(* Logix 5000 project; controller TFF vendor 1 type 14 code 107 rev 34.11; software revision 34.03; part 16 of 36 *)
(* tags used below, declared in another part *)
   Index : DINT;   // Index
   PLCDST : SINT;   // Current PLC Day Light Saving
   PLCTimeZoneString : STRING;   // Current PLC TimeZone
   TimeZoneUTC0 : STRING;   // String value for Time zone UTC 0
   Concentration : Concentration;
   ControlLoop_PCV001 : ALIAS FOR ControlLoop[3];   // PCV001 Control Loop
   ControlLoop_PCV001_5ms : ALIAS FOR ControlLoop[4];   // PCV001 Control Loop
   ControlLoop_PCV001_RAMP_OUT : REAL;   // Ramp Output
   Diafiltration : Diafiltration;
   FI101 : ALIAS FOR AnalogPoint[2];   // Filtrate Flow
   FQ_Conc : ALIAS FOR Totalizer[0];   // Concentration Totalizer
   FQ_Diaf : ALIAS FOR Totalizer[1];   // DiafiltrationTotalizer
   PCDateTime : DINT[7];   // Date/Time Array from PC
   PCV001 : ALIAS FOR AnalogPoint[3];   // Retentate Pressure Control Valve Position
   PCV001_Control : PCV_Control;   // PCV001 Control UDT
   PCV001_PID : PCV;   // PCV001 PID Management
   Phase : Phases[6];   // Phase Control Array
   PhaseTotalizer : PhaseTotalizer[18];   // Phase Totalizers Array
   Rack_Murr_Node1_TF2S : IO_Station;   // Status of Node 1 TF2S
   Rack_Murr_Node1_TF3S : IO_Station;   // Status of Node 1 TF3S
   RawAnalogInputArray : INT[50];   // Array of analog input raw
   SysControl : SysControl;   // General system status and command
   ThisSystem : SystemType;
   TimerControl : TimerControl;   // Timer Control
   Timers : Timers[22];   // Timer Array
   Totalizer : Totalizers[20];   // Totalizers Array
   Valve : Valve[100];   // Valve Array
(* MainProgram, continued *)

ROUTINE modTotal   (* ladder *)
// Totalizer Module
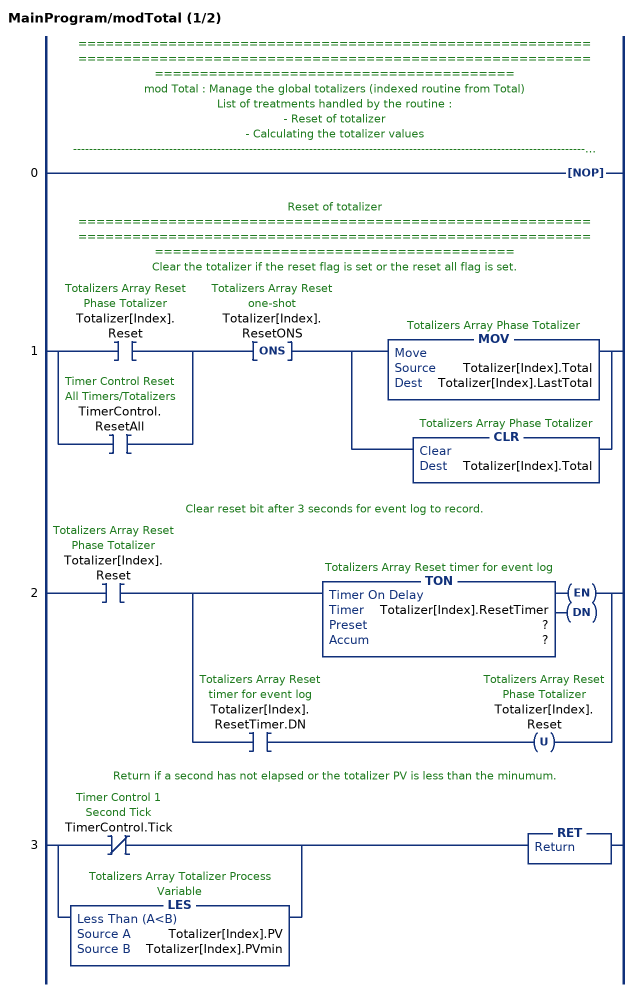
   // ==========================================================================================================================================================
   //                                                                                                   mod Total : Manage the global totalizers (indexed routine from Total)
   //                                                     List of treatments handled by the routine :
   //                                                          - Reset of totalizer
   //                                                          - Calculating the totalizer values
   //                                                     -----------------------------------------------------------------------------------------------------------------------------------------------------
   //                                                     History
   //                                                         2019-AUG-13 - Actemium - B. Roch - Initial version for Candidate Release 3.00.00.00.a
   // ==========================================================================================================================================================
   0: NOP();
   // Reset of totalizer
   // ==========================================================================================================================================================
   // Clear the totalizer if the reset flag is set or the reset all flag is set.
   1: [XIC(Totalizer[Index].Reset) ,XIC(TimerControl.ResetAll) ]ONS(Totalizer[Index].ResetONS)[MOV(Totalizer[Index].Total,Totalizer[Index].LastTotal) ,CLR(Totalizer[Index].Total) ];
   // Clear reset bit after 3 seconds for event log to record.
   2: XIC(Totalizer[Index].Reset)[TON(Totalizer[Index].ResetTimer,?,?) ,XIC(Totalizer[Index].ResetTimer.DN) OTU(Totalizer[Index].Reset) ];
   // Return if a second has not elapsed or the totalizer PV is less than the minumum.
   3: [XIO(TimerControl.Tick) ,LES(Totalizer[Index].PV,Totalizer[Index].PVmin) ]RET();
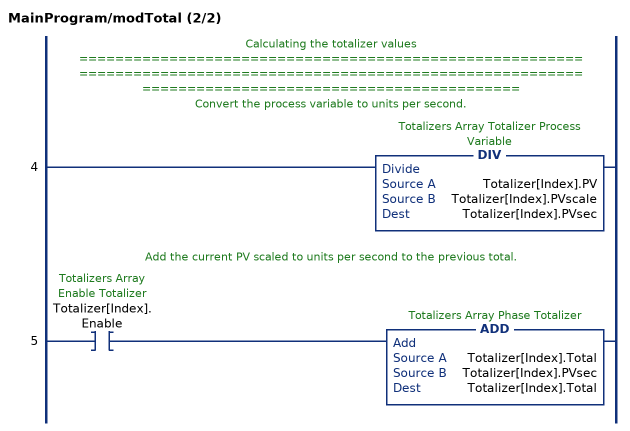
   // Calculating the totalizer values
   // ==========================================================================================================================================================
   // Convert the process variable to units per second.
   4: DIV(Totalizer[Index].PV,Totalizer[Index].PVscale,Totalizer[Index].PVsec);
   // Add the current PV scaled to units per second to the previous total.
   5: XIC(Totalizer[Index].Enable)ADD(Totalizer[Index].Total,Totalizer[Index].PVsec,Totalizer[Index].Total);
END_ROUTINE

ROUTINE PCDateTime   (* structured text *)
   (* =======================================================================
   	PCDateTime : Synchronize the PLC with PC clock
   
   	List of treatments
   		- Synchronization
   
   -----------------------------------------------------------------------------------------------------------------------------------------------------
   	History
   		2019-AUG-13 - ACTEMIUM - B. Roch - Initial version for Candidate Release 3.00.00.00.a
   		2020-SEP-14 - MERCK - Q. Spindler - Modifications for Candidate Release 3.00.00.01.a
   					- Add PLC TimeZone and DST forced settings
   =========================================================================*)
   
   
   (* Synchronization
   =========================================================================*)
   (*Update the internal PLC clock with the PC clock when the microseconds value is not -1*)
   IF PCDateTime[6] <> -1 THEN;
   	SSV (WALLCLOCKTIME, , DateTime, PCDateTime[0]);
   	PCDateTime[6] := -1;
   END_IF;
   
   (*Get PLC DST settings and set it to 0 of not already*)
   GSV (WALLCLOCKTIME, ,ApplyDST , PLCDST);
   IF PLCDST <> 0 THEN;
   	PLCDST := 0;
   	SSV (WALLCLOCKTIME, ,ApplyDST , PLCDST);
   END_IF;
   
   (*Get PLC TimeZone and set it to UTC0 of not already*)
   GSV (WALLCLOCKTIME, ,TimeZoneString, PLCTimeZoneString);
   IF PLCTimeZoneString <> TimeZoneUTC0 THEN;
   	SSV (WALLCLOCKTIME, ,TimeZoneString , TimeZoneUTC0);
   END_IF;
   
END_ROUTINE

ROUTINE Time   (* ladder *)
// Timekeeping Routine
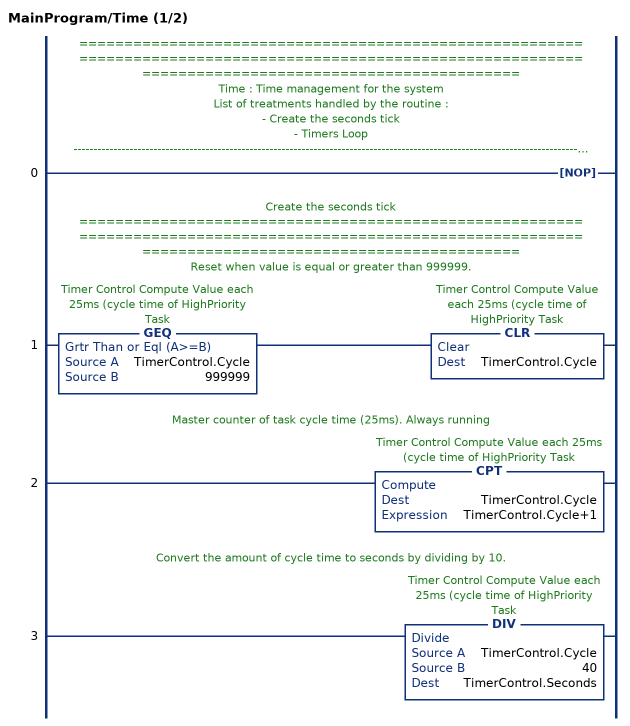
   // ==========================================================================================================================================================
   //                                                                                                                       Time : Time management for the system
   //                                                     List of treatments handled by the routine :
   //                                                          - Create the seconds tick
   //                                                          - Timers Loop
   //                                                     -----------------------------------------------------------------------------------------------------------------------------------------------------
   //                                                     History
   //                                                          2019-AUG-13 - Actemium - B. Roch - Initial version for Candidate Release 3.00.00.00.a
   //                                                          2020-SEP-14 - Merck - Q. Spindler - Modifications for Candidate Release 3.00.00.01.a
   //                                                                  - Add TimerControl.NewTickMainTask for 1 sec tick in Main task
   // ==========================================================================================================================================================
   0: NOP();
   // Create the seconds tick
   // ==========================================================================================================================================================
   // Reset when value is equal or greater than 999999.
   1: GEQ(TimerControl.Cycle,999999)CLR(TimerControl.Cycle);
   // Master counter of task cycle time (25ms). Always running
   2: CPT(TimerControl.Cycle,TimerControl.Cycle+1);
   // Convert the amount of cycle time to seconds by dividing by 10.
   3: DIV(TimerControl.Cycle,40,TimerControl.Seconds);
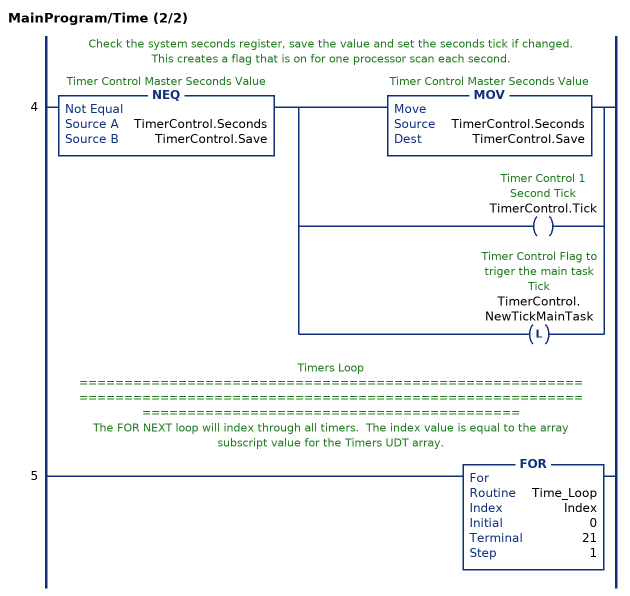
   // Check the system seconds register, save the value and set the seconds tick if changed.  This creates a flag that is on for one processor scan each second.
   4: NEQ(TimerControl.Seconds,TimerControl.Save)[MOV(TimerControl.Seconds,TimerControl.Save) ,OTE(TimerControl.Tick) ,OTL(TimerControl.NewTickMainTask) ];
   // Timers Loop
   // ==========================================================================================================================================================
   // The FOR NEXT loop will index through all timers.  The index value is equal to the array subscript value for the Timers UDT array.
   5: FOR(Time_Loop,Index,0,21,1);
END_ROUTINE

ROUTINE Time_Loop   (* ladder *)
// Timer Routine
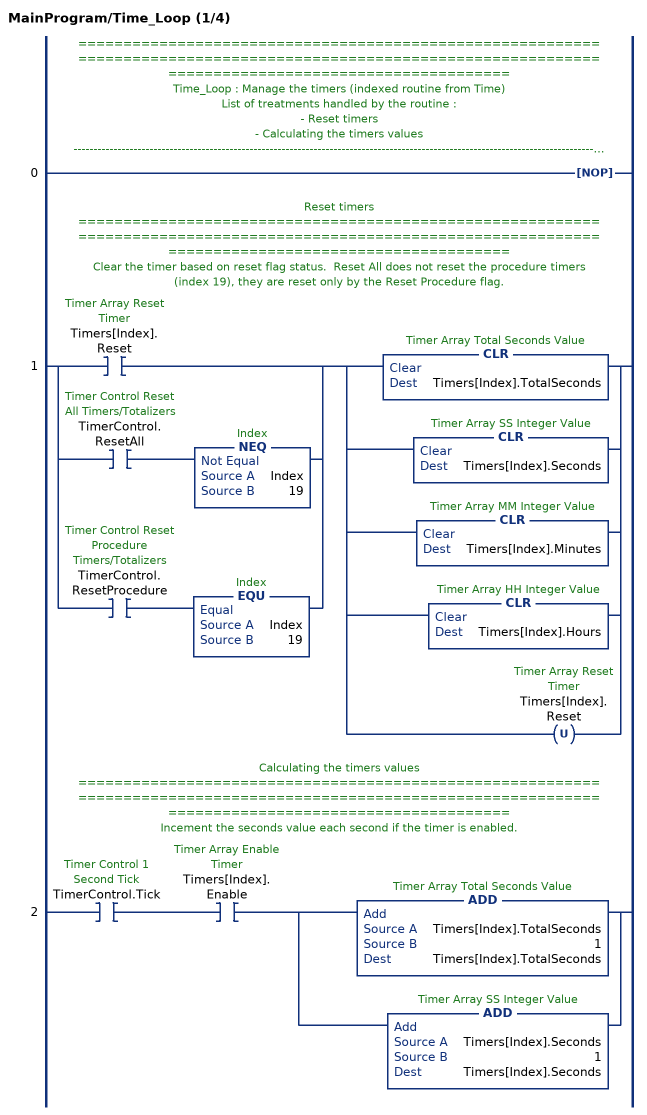
   // ==========================================================================================================================================================
   //                                                                                                              Time_Loop : Manage the timers (indexed routine from Time)
   //                                                     List of treatments handled by the routine :
   //                                                          - Reset timers
   //                                                          - Calculating the timers values
   //                                                     -----------------------------------------------------------------------------------------------------------------------------------------------------
   //                                                     History
   //                                                         2019-AUG-13 - Actemium - B. Roch - Initial version for Candidate Release 3.00.00.00.a
   // ==========================================================================================================================================================
   0: NOP();
   // Reset timers
   // ==========================================================================================================================================================
   // Clear the timer based on reset flag status.  Reset All does not reset the procedure timers (index 19), they are reset only by the Reset Procedure flag.
   1: [XIC(Timers[Index].Reset) ,XIC(TimerControl.ResetAll) NEQ(Index,19) ,XIC(TimerControl.ResetProcedure) EQU(Index,19) ][CLR(Timers[Index].TotalSeconds) ,CLR(Timers[Index].Seconds) ,CLR(Timers[Index].Minutes) ,CLR(Timers[Index].Hours) ,OTU(Timers[Index].Reset) ];
   // Calculating the timers values
   // ==========================================================================================================================================================
   // Incement the seconds value each second if the timer is enabled.
   2: XIC(TimerControl.Tick)XIC(Timers[Index].Enable)[ADD(Timers[Index].TotalSeconds,1,Timers[Index].TotalSeconds) ,ADD(Timers[Index].Seconds,1,Timers[Index].Seconds) ];
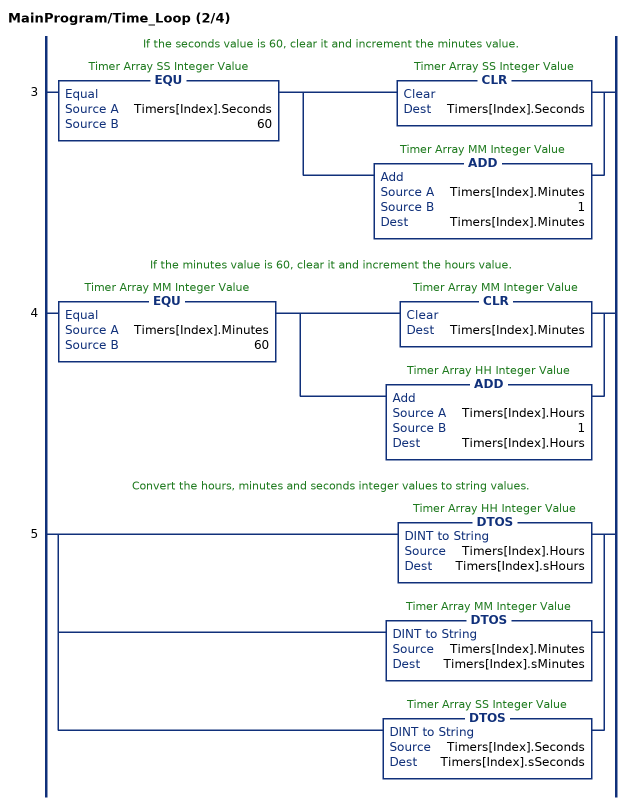
   // If the seconds value is 60, clear it and increment the minutes value.
   3: EQU(Timers[Index].Seconds,60)[CLR(Timers[Index].Seconds) ,ADD(Timers[Index].Minutes,1,Timers[Index].Minutes) ];
   // If the minutes value is 60, clear it and increment the hours value.
   4: EQU(Timers[Index].Minutes,60)[CLR(Timers[Index].Minutes) ,ADD(Timers[Index].Hours,1,Timers[Index].Hours) ];
   // Convert the hours, minutes and seconds integer values to string values.
   5: [DTOS(Timers[Index].Hours,Timers[Index].sHours) ,DTOS(Timers[Index].Minutes,Timers[Index].sMinutes) ,DTOS(Timers[Index].Seconds,Timers[Index].sSeconds) ];
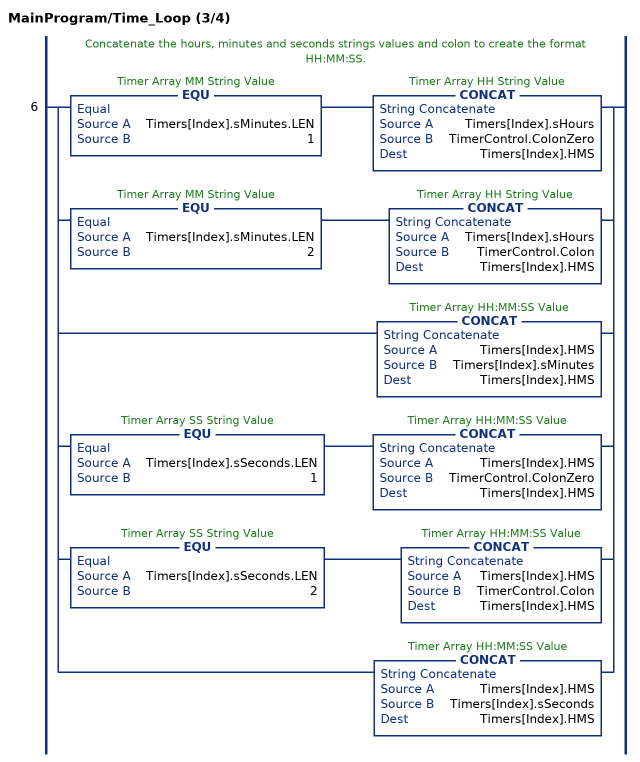
   // Concatenate the hours, minutes and seconds strings values and colon to create the format HH:MM:SS.
   6: [EQU(Timers[Index].sMinutes.LEN,1) CONCAT(Timers[Index].sHours,TimerControl.ColonZero,Timers[Index].HMS) ,EQU(Timers[Index].sMinutes.LEN,2) CONCAT(Timers[Index].sHours,TimerControl.Colon,Timers[Index].HMS) ,CONCAT(Timers[Index].HMS,Timers[Index].sMinutes,Timers[Index].HMS) ,EQU(Timers[Index].sSeconds.LEN,1) CONCAT(Timers[Index].HMS,TimerControl.ColonZero,Timers[Index].HMS) ,EQU(Timers[Index].sSeconds.LEN,2) CONCAT(Timers[Index].HMS,TimerControl.Colon,Timers[Index].HMS) ,CONCAT(Timers[Index].HMS,Timers[Index].sSeconds,Timers[Index].HMS) ];
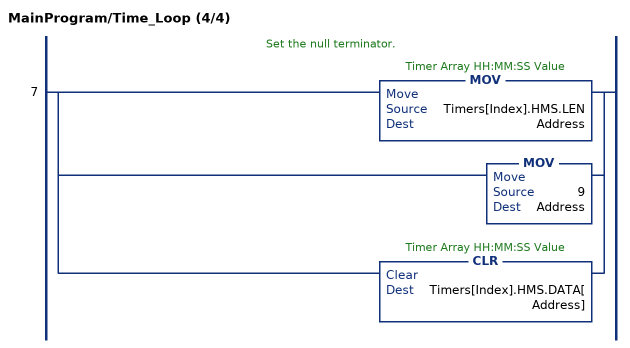
   // Set the null terminator.
   7: [[MOV(Timers[Index].HMS.LEN,Address) ,MOV(9,Address) ] ,CLR(Timers[Index].HMS.DATA[Address]) ];
END_ROUTINE

ROUTINE Total   (* ladder *)
// Totalizer Routine
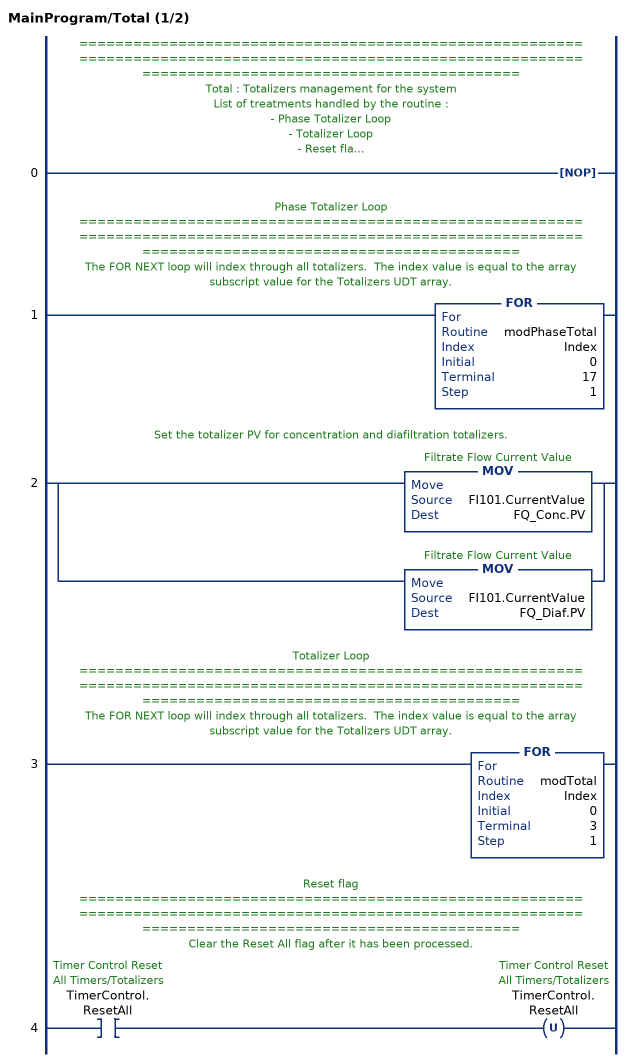
   // ==========================================================================================================================================================
   //                                                                                                              Total : Totalizers management for the system
   //                                                     List of treatments handled by the routine :
   //                                                          - Phase Totalizer Loop
   //                                                          - Totalizer Loop
   //                                                          - Reset flag
   //                                                     -----------------------------------------------------------------------------------------------------------------------------------------------------
   //                                                     History
   //                                                          2019-AUG-13 - Actemium - B. Roch - Initial version for Candidate Release 3.00.00.00.a
   // 		2020-SEP-29 - Merck - Q. Spindler - Modifications for Candidate Release 3.00.00.01.a
   // 							- Change array size of PhaseTotalizer
   // ==========================================================================================================================================================
   0: NOP();
   // Phase Totalizer Loop
   // ==========================================================================================================================================================
   // The FOR NEXT loop will index through all totalizers.  The index value is equal to the array subscript value for the Totalizers UDT array.
   1: FOR(modPhaseTotal,Index,0,17,1);
   // Set the totalizer PV for concentration and diafiltration totalizers.
   2: [MOV(FI101.CurrentValue,FQ_Conc.PV) ,MOV(FI101.CurrentValue,FQ_Diaf.PV) ];
   // Totalizer Loop
   // ==========================================================================================================================================================
   // The FOR NEXT loop will index through all totalizers.  The index value is equal to the array subscript value for the Totalizers UDT array.
   3: FOR(modTotal,Index,0,3,1);
   // Reset flag
   // ==========================================================================================================================================================
   // Clear the Reset All flag after it has been processed.
   4: XIC(TimerControl.ResetAll)OTU(TimerControl.ResetAll);
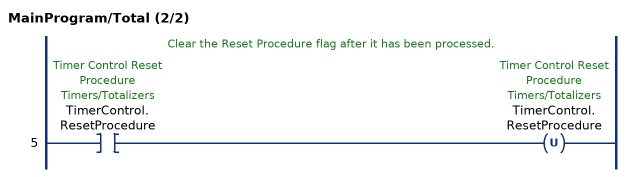
   // Clear the Reset Procedure flag after it has been processed.
   5: XIC(TimerControl.ResetProcedure)OTU(TimerControl.ResetProcedure);
END_ROUTINE
END_PROGRAM

PROGRAM MainProgram5ms   (* main routine MainRoutine, fault routine FaultRoutine *)
VAR
   Address : DINT := 1;   // Index
   Address2 : DINT := 41;
   ONS_PID02 : BOOL;
   PCV001_PID_Settings : INT;
   PCV101_PID_Settings : INT;
   SCL : SCALE := (InRawMax := 99999.0, InEUMax := 999.99);   // Scale Function
END_VAR

ROUTINE Control_Loop_PCV001_5ms   (* ladder *)
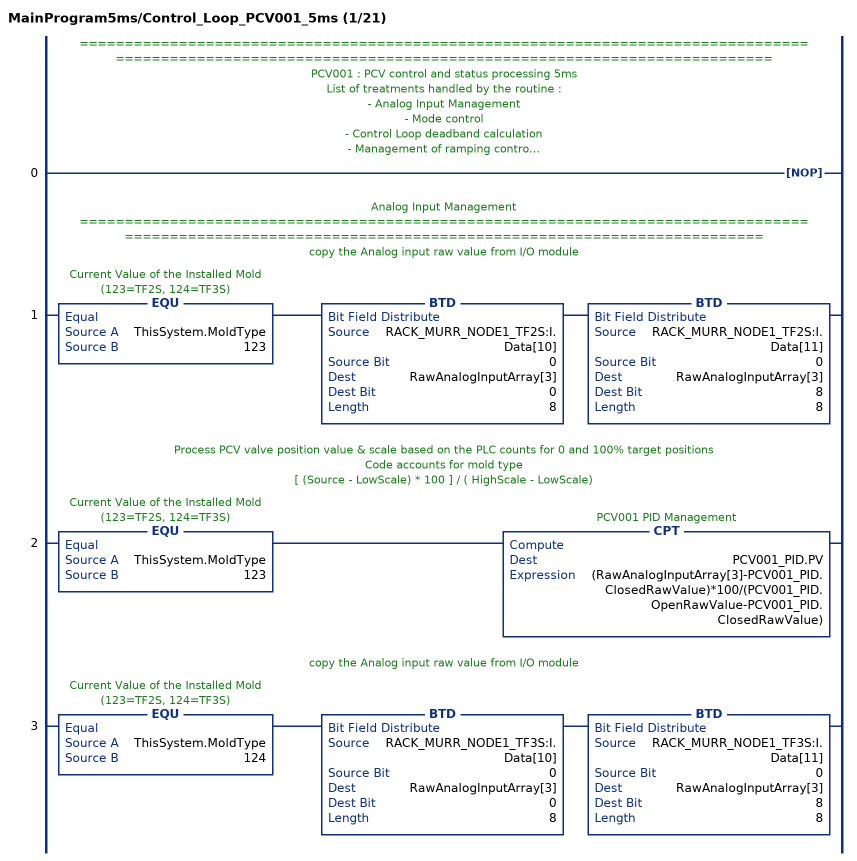
   // ==========================================================================================================================================================
   //                                                  PCV001 : PCV control and status processing 5ms
   //                                                     List of treatments handled by the routine :
   //                                                          - Analog Input Management
   //                                                          - Mode control
   //                                                          - Control Loop deadband calculation
   //                                                          - Management of ramping control
   //                                                          - Management of PID instruction
   //                                                          - PCV001 Control Valve Calibration
   //                                                          - Control of the analog output
   //                                                          - Loop status for HMI
   //                                                     -----------------------------------------------------------------------------------------------------------------------------------------------------
   //                                                     History
   //                                                          2019-AUG-13 - Actemium - B. Roch - Initial version for Candidate Release 3.00.00.00.a
   // 		                                2019-SEP-26 - ACTEMIUM - B. Roch - Modifications for Candidate Release 3.00.00.00.c
   // 					- Change compute for Analog Input Managment
   //                                                                                - Update Ramping up and down conditions
   // ==========================================================================================================================================================
   0: NOP();
   // Analog Input Management
   // ========================================================================================================================================================
   // copy the Analog input raw value from I/O module
   1: EQU(ThisSystem.MoldType,123)BTD(RACK_MURR_NODE1_TF2S:I.Data[10],0,RawAnalogInputArray[3],0,8)BTD(RACK_MURR_NODE1_TF2S:I.Data[11],0,RawAnalogInputArray[3],8,8);
   // Process PCV valve position value & scale based on the PLC counts for 0 and 100% target positions
   // Code accounts for mold type
   // [ (Source - LowScale) * 100 ] / ( HighScale - LowScale)
   2: EQU(ThisSystem.MoldType,123)CPT(PCV001_PID.PV,(RawAnalogInputArray[3]-PCV001_PID.ClosedRawValue)*100/(PCV001_PID.OpenRawValue-PCV001_PID.ClosedRawValue));
   // copy the Analog input raw value from I/O module
   3: EQU(ThisSystem.MoldType,124)BTD(RACK_MURR_NODE1_TF3S:I.Data[10],0,RawAnalogInputArray[3],0,8)BTD(RACK_MURR_NODE1_TF3S:I.Data[11],0,RawAnalogInputArray[3],8,8);
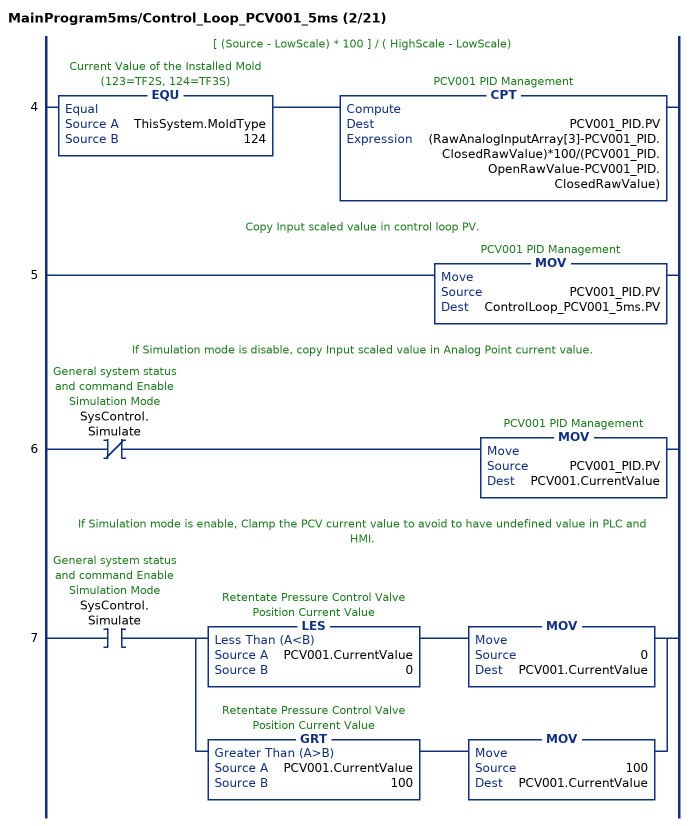
   // [ (Source - LowScale) * 100 ] / ( HighScale - LowScale)
   4: EQU(ThisSystem.MoldType,124)CPT(PCV001_PID.PV,(RawAnalogInputArray[3]-PCV001_PID.ClosedRawValue)*100/(PCV001_PID.OpenRawValue-PCV001_PID.ClosedRawValue));
   // Copy Input scaled value in control loop PV.
   5: MOV(PCV001_PID.PV,ControlLoop_PCV001_5ms.PV);
   // If Simulation mode is disable, copy Input scaled value in Analog Point current value.
   6: XIO(SysControl.Simulate)MOV(PCV001_PID.PV,PCV001.CurrentValue);
   // If Simulation mode is enable, Clamp the PCV current value to avoid to have undefined value in PLC and HMI.
   7: XIC(SysControl.Simulate)[LES(PCV001.CurrentValue,0) MOV(0,PCV001.CurrentValue) ,GRT(PCV001.CurrentValue,100) MOV(100,PCV001.CurrentValue) ];
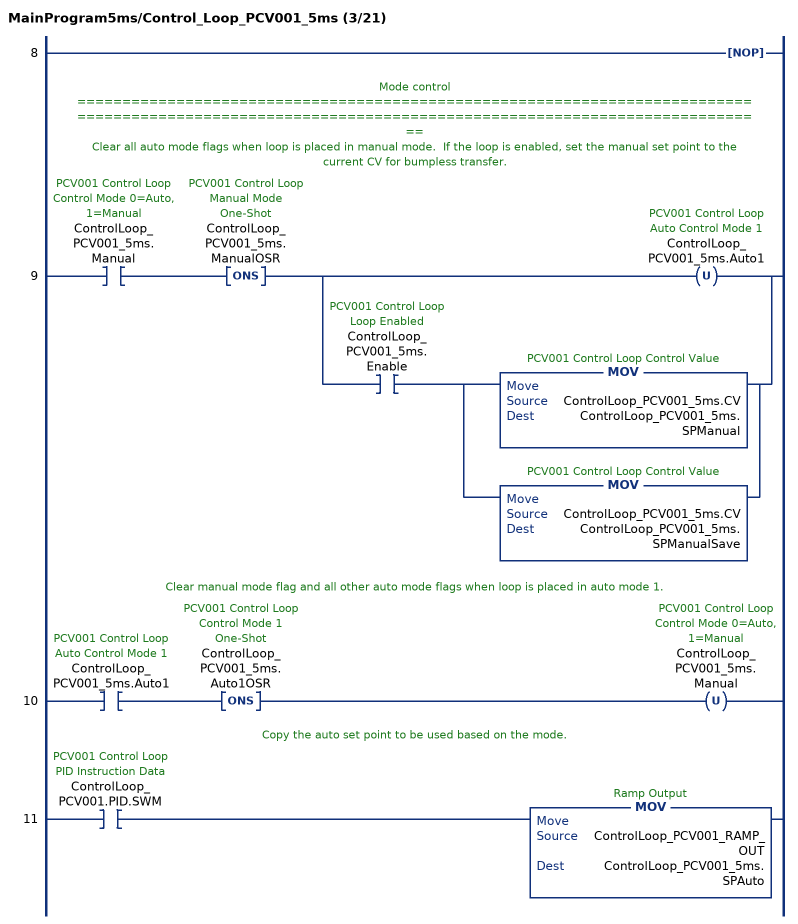
   8: NOP();
   // Mode control
   // ========================================================================================================================================================
   // Clear all auto mode flags when loop is placed in manual mode.  If the loop is enabled, set the manual set point to the current CV for bumpless transfer.
   9: XIC(ControlLoop_PCV001_5ms.Manual)ONS(ControlLoop_PCV001_5ms.ManualOSR)[OTU(ControlLoop_PCV001_5ms.Auto1) ,XIC(ControlLoop_PCV001_5ms.Enable) [MOV(ControlLoop_PCV001_5ms.CV,ControlLoop_PCV001_5ms.SPManual) ,MOV(ControlLoop_PCV001_5ms.CV,ControlLoop_PCV001_5ms.SPManualSave) ] ];
   // Clear manual mode flag and all other auto mode flags when loop is placed in auto mode 1.
   10: XIC(ControlLoop_PCV001_5ms.Auto1)ONS(ControlLoop_PCV001_5ms.Auto1OSR)OTU(ControlLoop_PCV001_5ms.Manual);
   // Copy the auto set point to be used based on the mode.
   11: XIC(ControlLoop_PCV001.PID.SWM)MOV(ControlLoop_PCV001_RAMP_OUT,ControlLoop_PCV001_5ms.SPAuto);
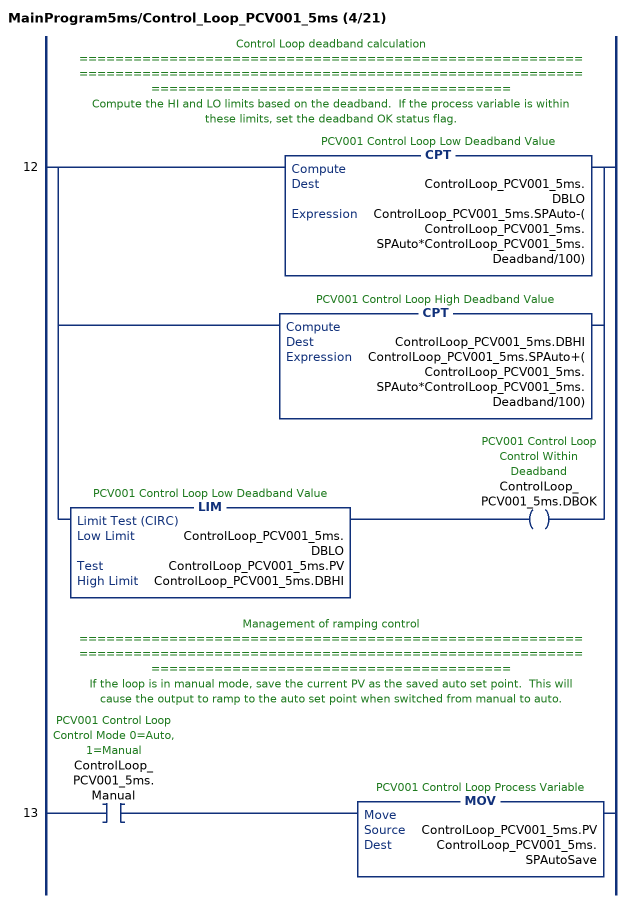
   // Control Loop deadband calculation
   // ========================================================================================================================================================
   // Compute the HI and LO limits based on the deadband.  If the process variable is within these limits, set the deadband OK status flag.
   12: [CPT(ControlLoop_PCV001_5ms.DBLO,ControlLoop_PCV001_5ms.SPAuto-(ControlLoop_PCV001_5ms.SPAuto*ControlLoop_PCV001_5ms.Deadband/100)) ,CPT(ControlLoop_PCV001_5ms.DBHI,ControlLoop_PCV001_5ms.SPAuto+(ControlLoop_PCV001_5ms.SPAuto*ControlLoop_PCV001_5ms.Deadband/100)) ,LIM(ControlLoop_PCV001_5ms.DBLO,ControlLoop_PCV001_5ms.PV,ControlLoop_PCV001_5ms.DBHI) OTE(ControlLoop_PCV001_5ms.DBOK) ];
   // Management of ramping control
   // ========================================================================================================================================================
   // If the loop is in manual mode, save the current PV as the saved auto set point.  This will cause the output to ramp to the auto set point when switched from manual to auto.
   13: XIC(ControlLoop_PCV001_5ms.Manual)MOV(ControlLoop_PCV001_5ms.PV,ControlLoop_PCV001_5ms.SPAutoSave);
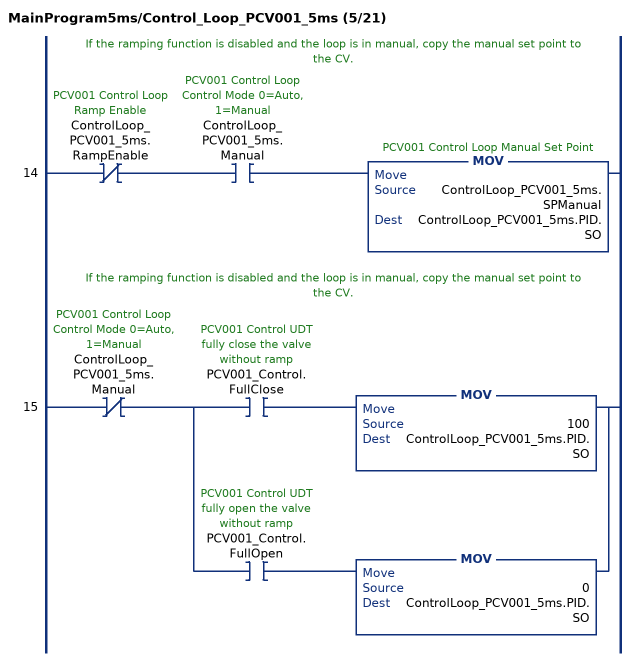
   // If the ramping function is disabled and the loop is in manual, copy the manual set point to the CV.
   14: XIO(ControlLoop_PCV001_5ms.RampEnable)XIC(ControlLoop_PCV001_5ms.Manual)MOV(ControlLoop_PCV001_5ms.SPManual,ControlLoop_PCV001_5ms.PID.SO);
   // If the ramping function is disabled and the loop is in manual, copy the manual set point to the CV.
   15: XIO(ControlLoop_PCV001_5ms.Manual)[XIC(PCV001_Control.FullClose) MOV(100,ControlLoop_PCV001_5ms.PID.SO) ,XIC(PCV001_Control.FullOpen) MOV(0,ControlLoop_PCV001_5ms.PID.SO) ];
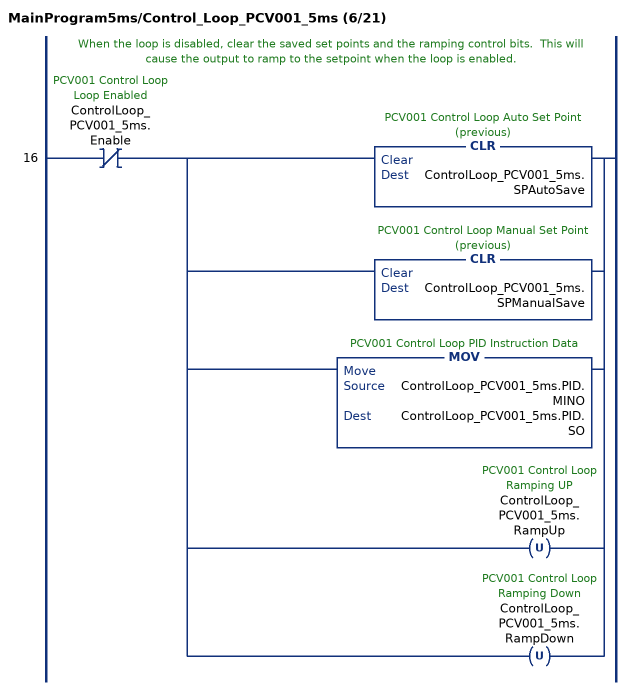
   // When the loop is disabled, clear the saved set points and the ramping control bits.  This will cause the output to ramp to the setpoint when the loop is enabled.
   16: XIO(ControlLoop_PCV001_5ms.Enable)[CLR(ControlLoop_PCV001_5ms.SPAutoSave) ,CLR(ControlLoop_PCV001_5ms.SPManualSave) ,MOV(ControlLoop_PCV001_5ms.PID.MINO,ControlLoop_PCV001_5ms.PID.SO) ,OTU(ControlLoop_PCV001_5ms.RampUp) ,OTU(ControlLoop_PCV001_5ms.RampDown) ];
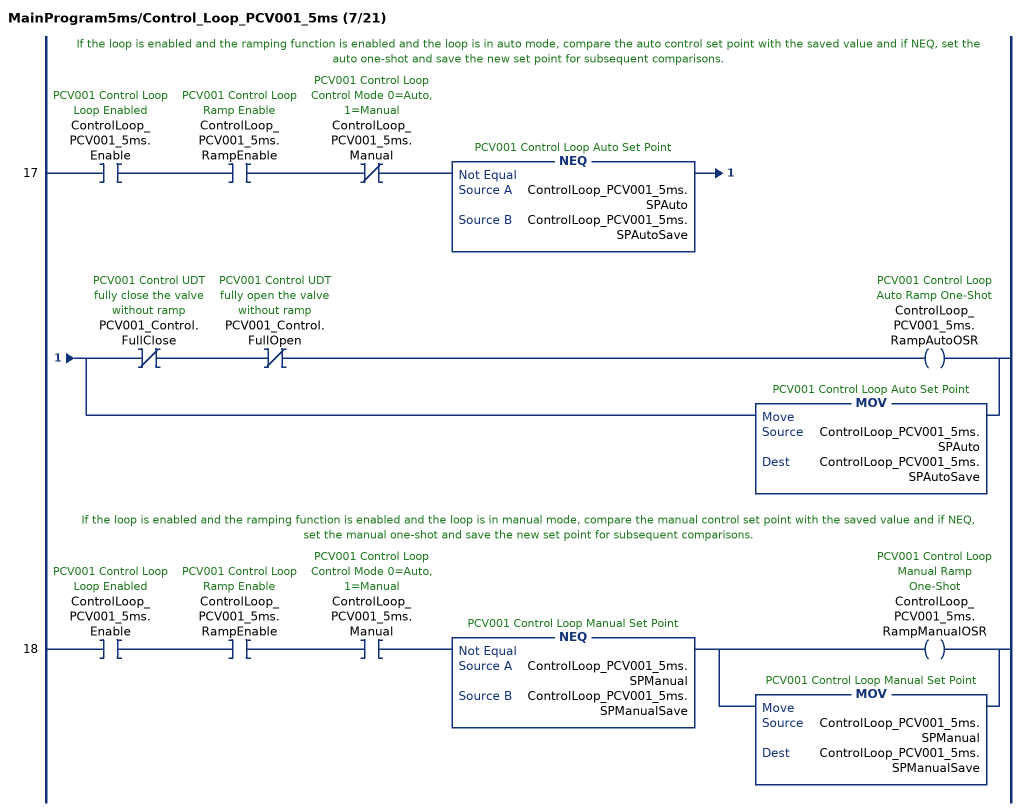
   // If the loop is enabled and the ramping function is enabled and the loop is in auto mode, compare the auto control set point with the saved value and if NEQ, set the auto one-shot and save the new set point for subsequent comparisons.
   17: XIC(ControlLoop_PCV001_5ms.Enable)XIC(ControlLoop_PCV001_5ms.RampEnable)XIO(ControlLoop_PCV001_5ms.Manual)NEQ(ControlLoop_PCV001_5ms.SPAuto,ControlLoop_PCV001_5ms.SPAutoSave)[XIO(PCV001_Control.FullClose) XIO(PCV001_Control.FullOpen) OTE(ControlLoop_PCV001_5ms.RampAutoOSR) ,MOV(ControlLoop_PCV001_5ms.SPAuto,ControlLoop_PCV001_5ms.SPAutoSave) ];
   // If the loop is enabled and the ramping function is enabled and the loop is in manual mode, compare the manual control set point with the saved value and if NEQ, set the manual one-shot and save the new set point for subsequent comparisons.
   18: XIC(ControlLoop_PCV001_5ms.Enable)XIC(ControlLoop_PCV001_5ms.RampEnable)XIC(ControlLoop_PCV001_5ms.Manual)NEQ(ControlLoop_PCV001_5ms.SPManual,ControlLoop_PCV001_5ms.SPManualSave)[OTE(ControlLoop_PCV001_5ms.RampManualOSR) ,MOV(ControlLoop_PCV001_5ms.SPManual,ControlLoop_PCV001_5ms.SPManualSave) ];
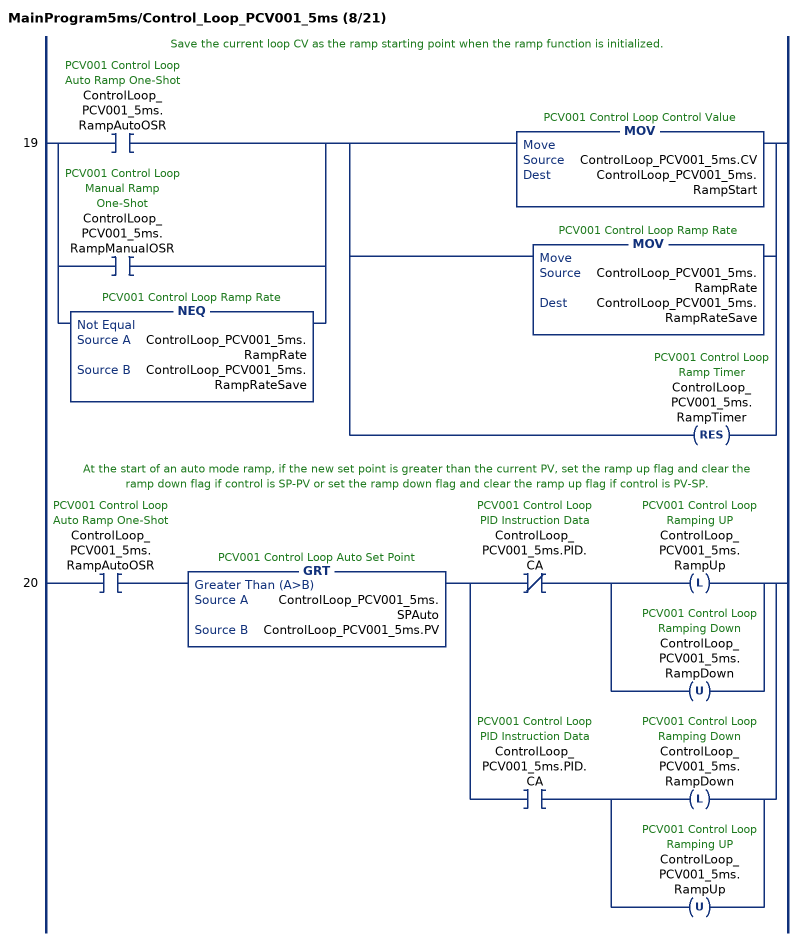
   // Save the current loop CV as the ramp starting point when the ramp function is initialized.
   19: [XIC(ControlLoop_PCV001_5ms.RampAutoOSR) ,XIC(ControlLoop_PCV001_5ms.RampManualOSR) ,NEQ(ControlLoop_PCV001_5ms.RampRate,ControlLoop_PCV001_5ms.RampRateSave) ][MOV(ControlLoop_PCV001_5ms.CV,ControlLoop_PCV001_5ms.RampStart) ,MOV(ControlLoop_PCV001_5ms.RampRate,ControlLoop_PCV001_5ms.RampRateSave) ,RES(ControlLoop_PCV001_5ms.RampTimer) ];
   // At the start of an auto mode ramp, if the new set point is greater than the current PV, set the ramp up flag and clear the ramp down flag if control is SP-PV or set the ramp down flag and clear the ramp up flag if control is PV-SP.
   20: XIC(ControlLoop_PCV001_5ms.RampAutoOSR)GRT(ControlLoop_PCV001_5ms.SPAuto,ControlLoop_PCV001_5ms.PV)[XIO(ControlLoop_PCV001_5ms.PID.CA) [OTL(ControlLoop_PCV001_5ms.RampUp) ,OTU(ControlLoop_PCV001_5ms.RampDown) ] ,XIC(ControlLoop_PCV001_5ms.PID.CA) [OTL(ControlLoop_PCV001_5ms.RampDown) ,OTU(ControlLoop_PCV001_5ms.RampUp) ] ];
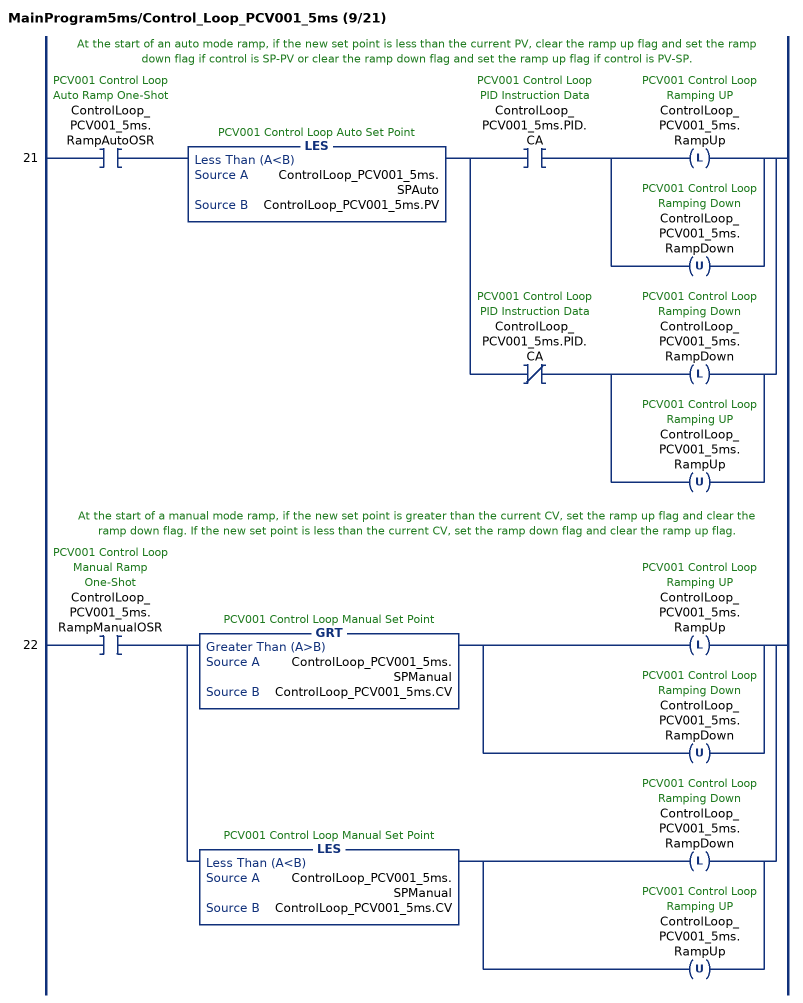
   // At the start of an auto mode ramp, if the new set point is less than the current PV, clear the ramp up flag and set the ramp down flag if control is SP-PV or clear the ramp down flag and set the ramp up flag if control is PV-SP.
   21: XIC(ControlLoop_PCV001_5ms.RampAutoOSR)LES(ControlLoop_PCV001_5ms.SPAuto,ControlLoop_PCV001_5ms.PV)[XIC(ControlLoop_PCV001_5ms.PID.CA) [OTL(ControlLoop_PCV001_5ms.RampUp) ,OTU(ControlLoop_PCV001_5ms.RampDown) ] ,XIO(ControlLoop_PCV001_5ms.PID.CA) [OTL(ControlLoop_PCV001_5ms.RampDown) ,OTU(ControlLoop_PCV001_5ms.RampUp) ] ];
   // At the start of a manual mode ramp, if the new set point is greater than the current CV, set the ramp up flag and clear the ramp down flag. If the new set point is less than the current CV, set the ramp down flag and clear the ramp up flag.
   22: XIC(ControlLoop_PCV001_5ms.RampManualOSR)[GRT(ControlLoop_PCV001_5ms.SPManual,ControlLoop_PCV001_5ms.CV) [OTL(ControlLoop_PCV001_5ms.RampUp) ,OTU(ControlLoop_PCV001_5ms.RampDown) ] ,LES(ControlLoop_PCV001_5ms.SPManual,ControlLoop_PCV001_5ms.CV) [OTL(ControlLoop_PCV001_5ms.RampDown) ,OTU(ControlLoop_PCV001_5ms.RampUp) ] ];
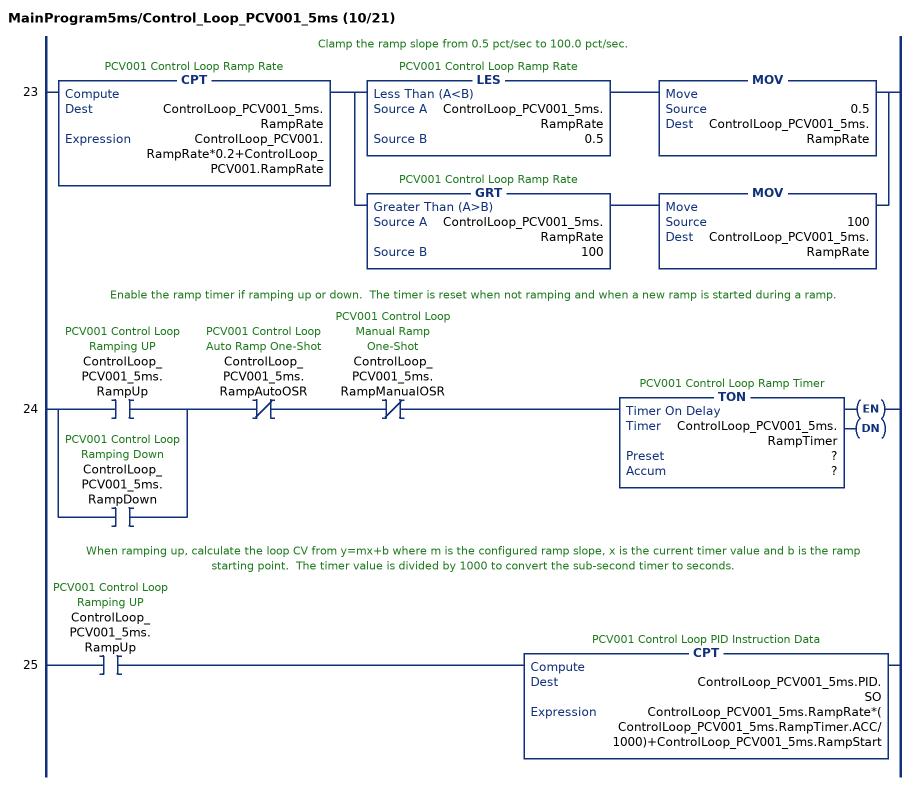
   // Clamp the ramp slope from 0.5 pct/sec to 100.0 pct/sec.
   23: CPT(ControlLoop_PCV001_5ms.RampRate,ControlLoop_PCV001.RampRate*0.2+ControlLoop_PCV001.RampRate)[LES(ControlLoop_PCV001_5ms.RampRate,0.5) MOV(0.5,ControlLoop_PCV001_5ms.RampRate) ,GRT(ControlLoop_PCV001_5ms.RampRate,100) MOV(100,ControlLoop_PCV001_5ms.RampRate) ];
   // Enable the ramp timer if ramping up or down.  The timer is reset when not ramping and when a new ramp is started during a ramp.
   24: [XIC(ControlLoop_PCV001_5ms.RampUp) ,XIC(ControlLoop_PCV001_5ms.RampDown) ]XIO(ControlLoop_PCV001_5ms.RampAutoOSR)XIO(ControlLoop_PCV001_5ms.RampManualOSR)TON(ControlLoop_PCV001_5ms.RampTimer,?,?);
   // When ramping up, calculate the loop CV from y=mx+b where m is the configured ramp slope, x is the current timer value and b is the ramp starting point.  The timer value is divided by 1000 to convert the sub-second timer to seconds.
   25: XIC(ControlLoop_PCV001_5ms.RampUp)CPT(ControlLoop_PCV001_5ms.PID.SO,ControlLoop_PCV001_5ms.RampRate*(ControlLoop_PCV001_5ms.RampTimer.ACC/1000)+ControlLoop_PCV001_5ms.RampStart);
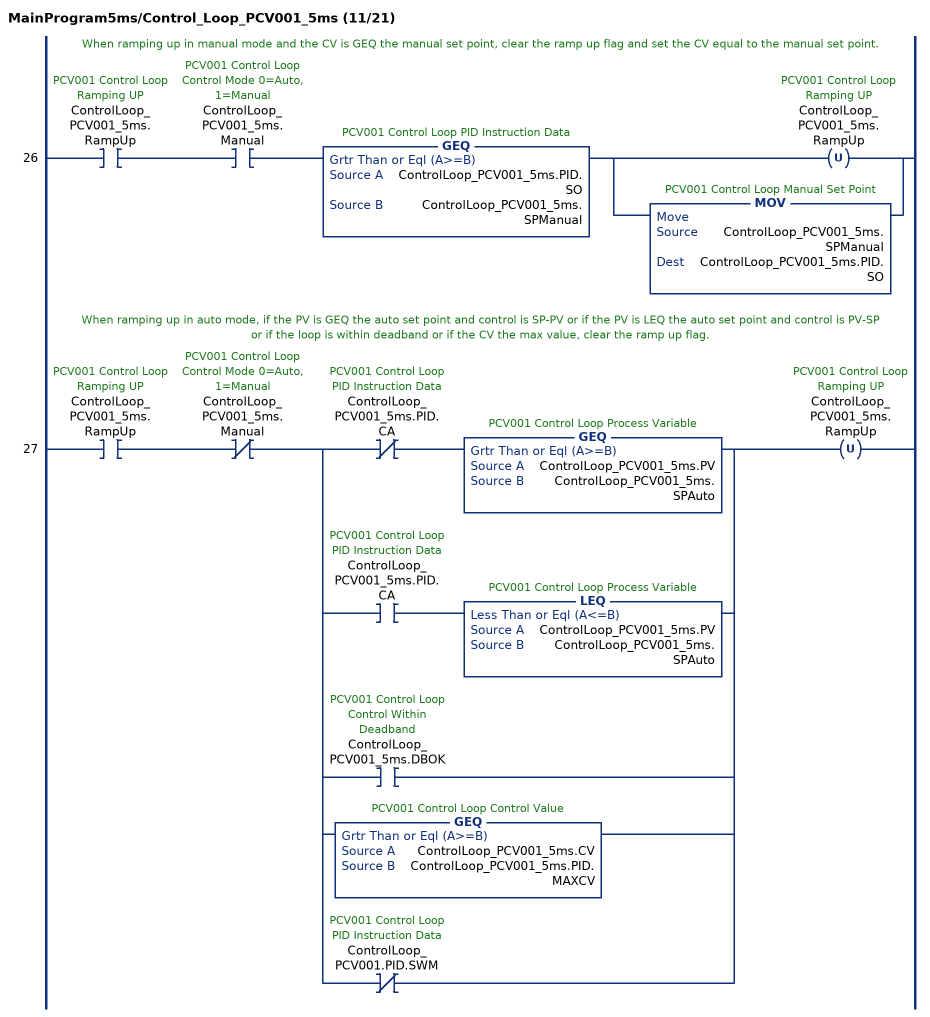
   // When ramping up in manual mode and the CV is GEQ the manual set point, clear the ramp up flag and set the CV equal to the manual set point.
   26: XIC(ControlLoop_PCV001_5ms.RampUp)XIC(ControlLoop_PCV001_5ms.Manual)GEQ(ControlLoop_PCV001_5ms.PID.SO,ControlLoop_PCV001_5ms.SPManual)[OTU(ControlLoop_PCV001_5ms.RampUp) ,MOV(ControlLoop_PCV001_5ms.SPManual,ControlLoop_PCV001_5ms.PID.SO) ];
   // When ramping up in auto mode, if the PV is GEQ the auto set point and control is SP-PV or if the PV is LEQ the auto set point and control is PV-SP or if the loop is within deadband or if the CV the max value, clear the ramp up flag.
   27: XIC(ControlLoop_PCV001_5ms.RampUp)XIO(ControlLoop_PCV001_5ms.Manual)[XIO(ControlLoop_PCV001_5ms.PID.CA) GEQ(ControlLoop_PCV001_5ms.PV,ControlLoop_PCV001_5ms.SPAuto) ,XIC(ControlLoop_PCV001_5ms.PID.CA) LEQ(ControlLoop_PCV001_5ms.PV,ControlLoop_PCV001_5ms.SPAuto) ,XIC(ControlLoop_PCV001_5ms.DBOK) ,[GEQ(ControlLoop_PCV001_5ms.CV,ControlLoop_PCV001_5ms.PID.MAXCV) ,XIO(ControlLoop_PCV001.PID.SWM) ] ]OTU(ControlLoop_PCV001_5ms.RampUp);
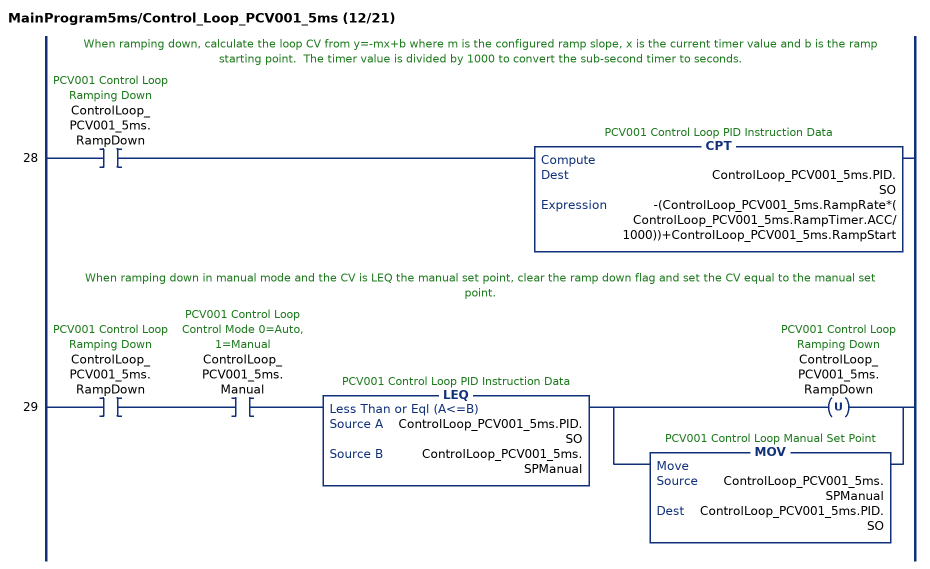
   // When ramping down, calculate the loop CV from y=-mx+b where m is the configured ramp slope, x is the current timer value and b is the ramp starting point.  The timer value is divided by 1000 to convert the sub-second timer to seconds.
   28: XIC(ControlLoop_PCV001_5ms.RampDown)CPT(ControlLoop_PCV001_5ms.PID.SO,-(ControlLoop_PCV001_5ms.RampRate*(ControlLoop_PCV001_5ms.RampTimer.ACC/1000))+ControlLoop_PCV001_5ms.RampStart);
   // When ramping down in manual mode and the CV is LEQ the manual set point, clear the ramp down flag and set the CV equal to the manual set point.
   29: XIC(ControlLoop_PCV001_5ms.RampDown)XIC(ControlLoop_PCV001_5ms.Manual)LEQ(ControlLoop_PCV001_5ms.PID.SO,ControlLoop_PCV001_5ms.SPManual)[OTU(ControlLoop_PCV001_5ms.RampDown) ,MOV(ControlLoop_PCV001_5ms.SPManual,ControlLoop_PCV001_5ms.PID.SO) ];
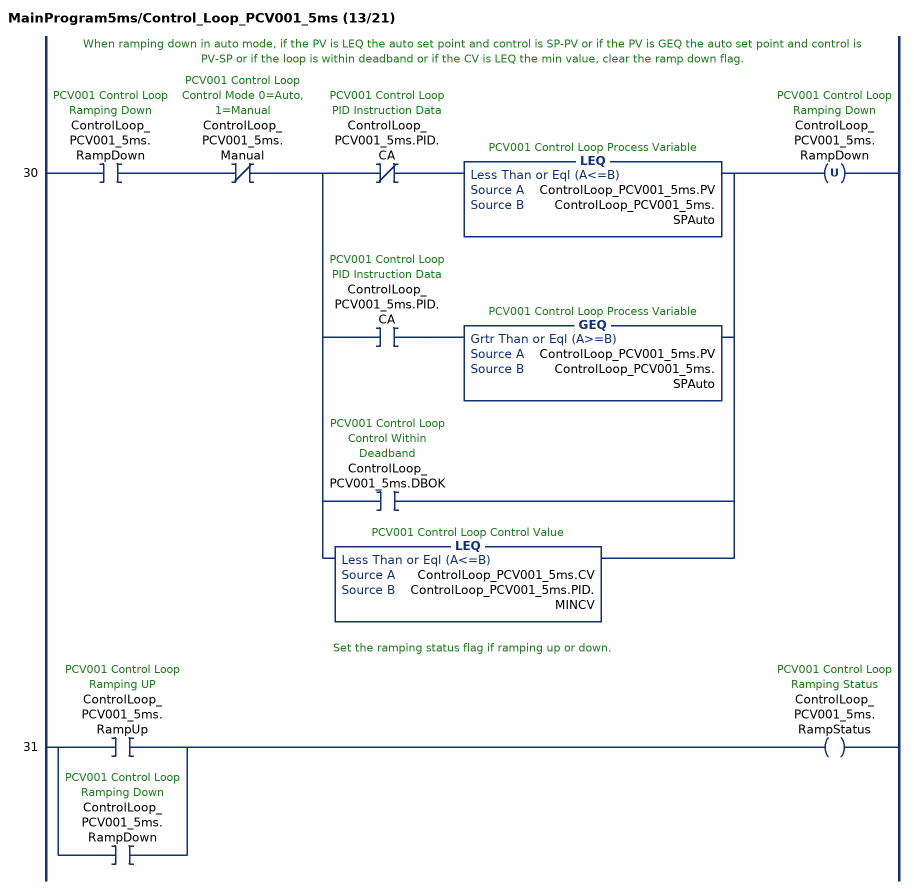
   // When ramping down in auto mode, if the PV is LEQ the auto set point and control is SP-PV or if the PV is GEQ the auto set point and control is PV-SP or if the loop is within deadband or if the CV is LEQ the min value, clear the ramp down flag.
   30: XIC(ControlLoop_PCV001_5ms.RampDown)XIO(ControlLoop_PCV001_5ms.Manual)[XIO(ControlLoop_PCV001_5ms.PID.CA) LEQ(ControlLoop_PCV001_5ms.PV,ControlLoop_PCV001_5ms.SPAuto) ,XIC(ControlLoop_PCV001_5ms.PID.CA) GEQ(ControlLoop_PCV001_5ms.PV,ControlLoop_PCV001_5ms.SPAuto) ,XIC(ControlLoop_PCV001_5ms.DBOK) ,LEQ(ControlLoop_PCV001_5ms.CV,ControlLoop_PCV001_5ms.PID.MINCV) ]OTU(ControlLoop_PCV001_5ms.RampDown);
   // Set the ramping status flag if ramping up or down.
   31: [XIC(ControlLoop_PCV001_5ms.RampUp) ,XIC(ControlLoop_PCV001_5ms.RampDown) ]OTE(ControlLoop_PCV001_5ms.RampStatus);
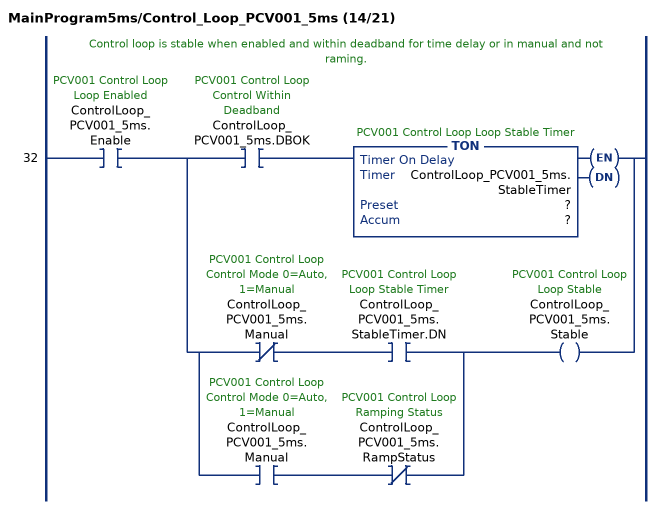
   // Control loop is stable when enabled and within deadband for time delay or in manual and not raming.
   32: XIC(ControlLoop_PCV001_5ms.Enable)[XIC(ControlLoop_PCV001_5ms.DBOK) TON(ControlLoop_PCV001_5ms.StableTimer,?,?) ,[XIO(ControlLoop_PCV001_5ms.Manual) XIC(ControlLoop_PCV001_5ms.StableTimer.DN) ,XIC(ControlLoop_PCV001_5ms.Manual) XIO(ControlLoop_PCV001_5ms.RampStatus) ] OTE(ControlLoop_PCV001_5ms.Stable) ];
